PROGRAM PRG_Chart
VAR
    bEnable, bIdle, bDone : BOOL;
    tonDelay : TON;
END_VAR

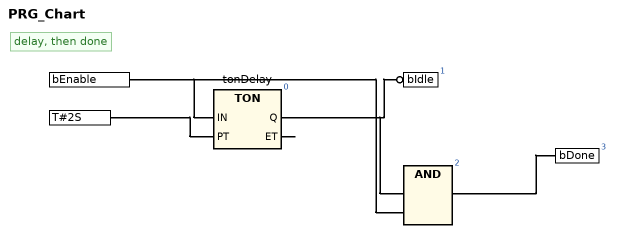
// delay, then done
tonDelay(IN := bEnable, PT := T#2S); // TON
bIdle := NOT tonDelay.Q;
bDone := tonDelay.Q AND bEnable;

END_PROGRAM

(* stored: Version 1.1.0.1, ProductVersion 3.1.4024.12
   POU PRG_Chart: Id {00000000-0000-0000-0000-000000000001}, SpecialFunc None *)
